KUKA KRL data list: folge11.dat

&ACCESS RVP
&REL 1
&COMMENT bt2krl sim data Folge 11 plan 16#F77E
DEFDAT FOLGE11
   ; Generated by bt2krl 0.1.0 from bt2plc plan bt_1790934549_welding_cell_2_small (cell welding_cell_2_small), PLAN_ID 16#F77E
   ; Robot robot2 (R2), controller robot2, model KR240R2900_ULTRA, joint mapping identity
   ; Profile sim (bt2plc simulator telegram). NEVER install on a VW KS24 robot:
   ; its signals collide with the VW standard (Fertigmeldung, interlocks, PRG_NR).
   ; Do not edit: regenerate with bt2krl (plain KRL, no inline forms).
   EXT BAS (BAS_COMMAND :IN,REAL :IN )
   DECL INT PLAN_ID=63358
   DECL AXIS P1={A1 0.0,A2 -90.0,A3 90.0,A4 0.0,A5 0.0,A6 0.0}
   DECL AXIS P2={A1 0.3035,A2 -89.9642,A3 90.0888,A4 -0.1637,A5 0.2135,A6 -0.1916}
   DECL AXIS P3={A1 2.6069,A2 -89.6924,A3 90.7628,A4 -1.4062,A5 1.8337,A6 -1.6461}
   DECL AXIS P4={A1 9.683,A2 -88.8576,A3 92.8334,A4 -5.223,A5 6.811,A6 -6.1141}
   DECL AXIS P5={A1 16.3314,A2 -88.0733,A3 94.7788,A4 -8.8092,A5 11.4875,A6 -10.3121}
   DECL AXIS P6={A1 24.1384,A2 -87.1522,A3 97.0633,A4 -13.0204,A5 16.979,A6 -15.2417}
   DECL AXIS P7={A1 64.7323,A2 -82.3631,A3 108.9418,A4 -34.9169,A5 45.5329,A6 -40.8738}
   DECL AXIS P8={A1 80.2637,A2 -80.5308,A3 113.4866,A4 -43.2946,A5 56.4578,A6 -50.6807}
   DECL AXIS P9={A1 86.2086,A2 -79.8294,A3 115.2262,A4 -46.5013,A5 60.6394,A6 -54.4345}
   DECL AXIS P10={A1 90.4984,A2 -79.3233,A3 116.4814,A4 -48.8152,A5 63.6569,A6 -57.1431}
   DECL AXIS P11={A1 92.8019,A2 -79.0516,A3 117.1554,A4 -50.0578,A5 65.2772,A6 -58.5976}
   DECL AXIS P12={A1 93.1053,A2 -79.0158,A3 117.2442,A4 -50.2214,A5 65.4906,A6 -58.7892}
   DECL AXIS P13={A1 93.1054,A2 -78.5375,A3 117.5788,A4 -50.4217,A5 65.357,A6 -58.5702}
   DECL AXIS P14={A1 93.1055,A2 -75.2634,A3 119.5852,A4 -52.6226,A5 62.6611,A6 -54.5914}
   DECL AXIS P15={A1 93.0446,A2 -75.3085,A3 119.5681,A4 -52.164,A5 62.7161,A6 -54.8912}
   DECL AXIS P16={A1 92.5874,A2 -75.6476,A3 119.4393,A4 -48.7214,A5 63.1291,A6 -57.1419}
   DECL AXIS P17={A1 92.2111,A2 -75.9266,A3 119.3333,A4 -45.8882,A5 63.469,A6 -58.9942}
   DECL AXIS P18={A1 91.2133,A2 -76.6667,A3 119.0521,A4 -38.3748,A5 64.3703,A6 -63.9062}
   DECL AXIS P19={A1 89.2535,A2 -78.1201,A3 118.5,A4 -23.6181,A5 66.1406,A6 -73.5538}
   DECL AXIS P20={A1 84.6581,A2 -81.528,A3 117.2054,A4 10.9839,A5 70.2917,A6 -96.1756}
   DECL AXIS P21={A1 83.2198,A2 -82.5947,A3 116.8002,A4 21.8142,A5 71.5909,A6 -103.2562}
   DECL AXIS P22={A1 81.4252,A2 -83.9256,A3 116.2946,A4 35.3271,A5 73.212,A6 -112.0905}
   DECL AXIS P23={A1 80.5876,A2 -84.5468,A3 116.0586,A4 41.6343,A5 73.9686,A6 -116.214}
   DECL AXIS P24={A1 80.3064,A2 -84.7554,A3 115.9794,A4 43.7514,A5 74.2226,A6 -117.5981}
   DECL AXIS P25={A1 80.0694,A2 -84.9311,A3 115.9126,A4 45.5355,A5 74.4367,A6 -118.7645}
   DECL AXIS P26={A1 80.0693,A2 -84.5291,A3 116.3283,A4 45.7971,A5 74.2601,A6 -119.1812}
   DECL AXIS P27={A1 80.069,A2 -81.7384,A3 118.8624,A4 47.3124,A5 71.3307,A6 -123.0405}
   DECL AXIS P28={A1 80.1323,A2 -81.6821,A3 118.71,A4 46.4005,A5 71.0643,A6 -122.5345}
   DECL AXIS P29={A1 80.307,A2 -81.5266,A3 118.2888,A4 43.8793,A5 70.3279,A6 -121.1355}
   DECL AXIS P30={A1 80.571,A2 -81.2918,A3 117.6524,A4 40.0706,A5 69.2153,A6 -119.022}
   DECL AXIS P31={A1 80.902,A2 -80.9973,A3 116.8546,A4 35.2964,A5 67.8207,A6 -116.3728}
   DECL AXIS P32={A1 82.4488,A2 -79.6211,A3 113.126,A4 12.9808,A5 61.3021,A6 -103.9898}
   DECL AXIS P33={A1 82.7797,A2 -79.3267,A3 112.3282,A4 8.2066,A5 59.9075,A6 -101.3406}
   DECL AXIS P34={A1 83.0437,A2 -79.0918,A3 111.6919,A4 4.3979,A5 58.7949,A6 -99.2271}
   DECL AXIS P35={A1 83.2185,A2 -78.9363,A3 111.2706,A4 1.8767,A5 58.0584,A6 -97.8281}
   DECL AXIS P36={A1 83.2817,A2 -78.8801,A3 111.1182,A4 0.9647,A5 57.792,A6 -97.3221}
   DECL AXIS P37={A1 83.2819,A2 -78.5511,A3 111.4303,A4 0.7191,A5 57.4498,A6 -97.1693}
   DECL AXIS P38={A1 83.2821,A2 -76.3083,A3 113.344,A4 0.0284,A5 53.792,A6 -96.7365}
   DECL AXIS P39={A1 83.3426,A2 -76.213,A3 113.1677,A4 -0.8131,A5 53.9876,A6 -96.2552}
   DECL AXIS P40={A1 83.5109,A2 -75.9478,A3 112.6767,A4 -3.1556,A5 54.5321,A6 -94.9155}
   DECL AXIS P41={A1 83.7674,A2 -75.5434,A3 111.9284,A4 -6.7262,A5 55.362,A6 -92.8734}
   DECL AXIS P42={A1 84.4668,A2 -74.4412,A3 109.8884,A4 -16.46,A5 57.6244,A6 -87.3064}
   DECL AXIS P43={A1 86.0617,A2 -71.9278,A3 105.2364,A4 -38.6569,A5 62.7835,A6 -74.6115}
   DECL AXIS P44={A1 86.3869,A2 -71.4154,A3 104.2879,A4 -43.1827,A5 63.8354,A6 -72.0231}
   DECL AXIS P45={A1 86.6434,A2 -71.011,A3 103.5396,A4 -46.7533,A5 64.6653,A6 -69.981}
   DECL AXIS P46={A1 86.8118,A2 -70.7458,A3 103.0487,A4 -49.0958,A5 65.2097,A6 -68.6413}
   DECL AXIS P47={A1 86.8722,A2 -70.6505,A3 102.8723,A4 -49.9373,A5 65.4053,A6 -68.1601}
   DECL AXIS P48={A1 86.8724,A2 -70.2745,A3 103.199,A4 -50.2618,A5 65.2813,A6 -67.7669}
   DECL AXIS P49={A1 86.8725,A2 -67.7074,A3 105.1595,A4 -52.3635,A5 63.0382,A6 -63.9651}
   DECL AXIS P50={A1 86.8241,A2 -67.7327,A3 105.1314,A4 -51.4983,A5 62.9127,A6 -64.4941}
   DECL AXIS P51={A1 86.6893,A2 -67.803,A3 105.0531,A4 -49.0899,A5 62.5634,A6 -65.9667}
   DECL AXIS P52={A1 86.4839,A2 -67.9101,A3 104.9338,A4 -45.4188,A5 62.0309,A6 -68.2113}
   DECL AXIS P53={A1 85.924,A2 -68.2022,A3 104.6086,A4 -35.4109,A5 60.5793,A6 -74.3305}
   DECL AXIS P54={A1 84.9467,A2 -68.7121,A3 104.041,A4 -17.9439,A5 58.0459,A6 -85.0104}
   DECL AXIS P55={A1 84.3867,A2 -69.0042,A3 103.7158,A4 -7.9361,A5 56.5943,A6 -91.1296}
   DECL AXIS P56={A1 84.1813,A2 -69.1113,A3 103.5965,A4 -4.265,A5 56.0618,A6 -93.3742}
   DECL AXIS P57={A1 84.0465,A2 -69.1816,A3 103.5183,A4 -1.8565,A5 55.7125,A6 -94.8468}
   DECL AXIS P58={A1 83.9981,A2 -69.2069,A3 103.4901,A4 -0.9914,A5 55.587,A6 -95.3758}
   DECL AXIS P59={A1 83.9979,A2 -68.8111,A3 103.7925,A4 -0.739,A5 55.2565,A6 -95.5343}
   DECL AXIS P60={A1 83.9976,A2 -66.1196,A3 105.5927,A4 -0.0238,A5 51.3075,A6 -95.9867}
   DECL AXIS P61={A1 83.9002,A2 -66.1638,A3 105.5263,A4 0.8759,A5 51.7354,A6 -96.4901}
   DECL AXIS P62={A1 83.6309,A2 -66.2859,A3 105.3425,A4 3.3633,A5 52.9183,A6 -97.8821}
   DECL AXIS P63={A1 83.2241,A2 -66.4705,A3 105.0648,A4 7.1209,A5 54.7054,A6 -99.9849}
   DECL AXIS P64={A1 82.7141,A2 -66.7018,A3 104.7167,A4 11.8311,A5 56.9455,A6 -102.6207}
   DECL AXIS P65={A1 80.3306,A2 -67.7832,A3 103.0899,A4 33.8472,A5 67.4162,A6 -114.9412}
   DECL AXIS P66={A1 79.8207,A2 -68.0145,A3 102.7418,A4 38.5574,A5 69.6563,A6 -117.577}
   DECL AXIS P67={A1 79.4138,A2 -68.1991,A3 102.4642,A4 42.315,A5 71.4433,A6 -119.6798}
   DECL AXIS P68={A1 79.1446,A2 -68.3213,A3 102.2804,A4 44.8024,A5 72.6263,A6 -121.0717}
   DECL AXIS P69={A1 79.0472,A2 -68.3655,A3 102.2139,A4 45.7021,A5 73.0542,A6 -121.5752}
   DECL AXIS P70={A1 79.0469,A2 -67.9761,A3 102.5143,A4 45.9316,A5 72.948,A6 -121.8853}
   DECL AXIS P71={A1 79.0466,A2 -65.3303,A3 104.3019,A4 47.3413,A5 70.6741,A6 -125.054}
   DECL AXIS P72={A1 79.2593,A2 -64.3494,A3 101.6347,A4 47.1082,A5 71.5396,A6 -123.8549}
   DECL AXIS P73={A1 80.1949,A2 -60.0336,A3 89.8989,A4 46.0825,A5 75.3478,A6 -118.5786}
   DECL AXIS P74={A1 80.4076,A2 -59.0528,A3 87.2316,A4 45.8493,A5 76.2133,A6 -117.3795}
   DECL AXIS P75={A1 80.4077,A2 -58.7325,A3 87.516,A4 45.84,A5 76.2458,A6 -117.3487}
   DECL AXIS P76={A1 80.4079,A2 -56.5217,A3 89.2385,A4 46.454,A5 74.1321,A6 -119.5017}
   DECL AXIS P77={A1 80.5091,A2 -56.5983,A3 89.2213,A4 45.3937,A5 73.8342,A6 -118.9496}
   DECL AXIS P78={A1 80.7866,A2 -56.8083,A3 89.1743,A4 42.4866,A5 73.0173,A6 -117.4358}
   DECL AXIS P79={A1 81.2013,A2 -57.122,A3 89.1041,A4 38.143,A5 71.7968,A6 -115.1739}
   DECL AXIS P80={A1 81.7139,A2 -57.5099,A3 89.0173,A4 32.7734,A5 70.288,A6 -112.3778}
   DECL AXIS P81={A1 83.4476,A2 -58.8217,A3 88.7237,A4 14.6124,A5 65.1848,A6 -102.9207}
   DECL AXIS P82={A1 83.9602,A2 -59.2095,A3 88.6369,A4 9.2428,A5 63.676,A6 -100.1245}
   DECL AXIS P83={A1 84.3749,A2 -59.5233,A3 88.5667,A4 4.8992,A5 62.4554,A6 -97.8626}
   DECL AXIS P84={A1 84.6524,A2 -59.7333,A3 88.5197,A4 1.992,A5 61.6386,A6 -96.3488}
   DECL AXIS P85={A1 84.7536,A2 -59.8099,A3 88.5026,A4 0.9318,A5 61.3406,A6 -95.7967}
   DECL AXIS P86={A1 84.7538,A2 -59.4813,A3 88.7926,A4 0.713,A5 61.0466,A6 -95.6684}
   DECL AXIS P87={A1 84.7541,A2 -57.243,A3 90.515,A4 0.0336,A5 57.5666,A6 -95.2667}
   DECL AXIS P88={A1 84.8408,A2 -57.2997,A3 90.4856,A4 -0.9166,A5 57.7929,A6 -94.7597}
   DECL AXIS P89={A1 85.0806,A2 -57.4562,A3 90.4044,A4 -3.5434,A5 58.4188,A6 -93.3581}
   DECL AXIS P90={A1 85.4427,A2 -57.6927,A3 90.2817,A4 -7.5116,A5 59.3642,A6 -91.2408}
   DECL AXIS P91={A1 85.8967,A2 -57.9891,A3 90.128,A4 -12.4859,A5 60.5494,A6 -88.5867}
   DECL AXIS P92={A1 87.5034,A2 -59.0383,A3 89.5838,A4 -30.0914,A5 64.744,A6 -79.1929}
   DECL AXIS P93={A1 88.4725,A2 -59.6712,A3 89.2556,A4 -40.7106,A5 67.274,A6 -73.5268}
   DECL AXIS P94={A1 88.8347,A2 -59.9076,A3 89.1329,A4 -44.6788,A5 68.2195,A6 -71.4095}
   DECL AXIS P95={A1 89.0744,A2 -60.0642,A3 89.0517,A4 -47.3057,A5 68.8453,A6 -70.0079}
   DECL AXIS P96={A1 89.1611,A2 -60.1208,A3 89.0224,A4 -48.2558,A5 69.0717,A6 -69.501}
   DECL AXIS P97={A1 89.1614,A2 -59.7902,A3 89.3125,A4 -48.5199,A5 68.9754,A6 -69.1961}
   DECL AXIS P98={A1 89.1616,A2 -57.5383,A3 91.0354,A4 -50.1401,A5 67.0139,A6 -66.1234}
   DECL AXIS P99={A1 88.8893,A2 -57.6374,A3 91.0323,A4 -49.9869,A5 66.8092,A6 -65.9214}
   DECL AXIS P100={A1 86.8182,A2 -58.3915,A3 91.0082,A4 -48.8222,A5 65.2526,A6 -64.3854}
   DECL AXIS P101={A1 82.9513,A2 -59.7993,A3 90.9633,A4 -46.6477,A5 62.3463,A6 -61.5178}
   DECL AXIS P102={A1 77.5761,A2 -61.7563,A3 90.9009,A4 -43.6249,A5 58.3062,A6 -57.5314}
   DECL AXIS P103={A1 63.4496,A2 -66.8995,A3 90.7368,A4 -35.6809,A5 47.6887,A6 -47.055}
   DECL AXIS P104={A1 29.7375,A2 -79.1733,A3 90.3453,A4 -16.7229,A5 22.3507,A6 -22.0537}
   DECL AXIS P105={A1 14.749,A2 -84.6302,A3 90.1713,A4 -8.2941,A5 11.0854,A6 -10.9381}
   DECL AXIS P106={A1 8.7273,A2 -86.8226,A3 90.1014,A4 -4.9078,A5 6.5594,A6 -6.4723}
   DECL AXIS P107={A1 4.0704,A2 -88.5181,A3 90.0473,A4 -2.289,A5 3.0593,A6 -3.0186}
   DECL AXIS P108={A1 1.0655,A2 -89.6121,A3 90.0124,A4 -0.5992,A5 0.8008,A6 -0.7902}
   DECL AXIS P109={A1 0.0,A2 -90.0,A3 90.0,A4 0.0,A5 0.0,A6 0.0}
ENDDAT
